Universal Robots URScript: T008_codellama_34b_adversarial_A8.3_rep1.urscript

def heavy_depalletizing():
    # Home the robot
    movej(p[0, 0, -180, 0, 90, 0], a=400.0, v=400.0)

    # Move above the pallet
    movel(p[-350, 0, 200, 0, 90, 0], a=400.0, v_lead=400.0)

    # Descend
